Universal Robots URScript: letra_E.script

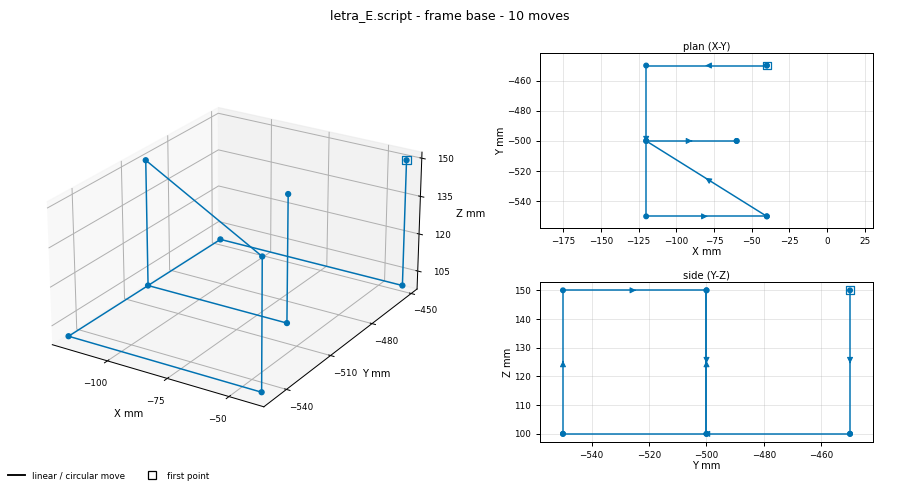
[picture p0: tool path of letra_E.script in frame base, 10 of 10 moves have a stored position in this frame; points joined in program order, loops and branches not executed]
# Letra E - Escobar
movel(p[-0.040, -0.450, 0.150, 3.1416, 0, 0], a=0.5, v=0.1)
movel(p[-0.040, -0.450, 0.100, 3.1416, 0, 0], a=0.5, v=0.1)
movel(p[-0.120, -0.450, 0.100, 3.1416, 0, 0], a=0.5, v=0.1)
movel(p[-0.120, -0.550, 0.100, 3.1416, 0, 0], a=0.5, v=0.1)
movel(p[-0.040, -0.550, 0.100, 3.1416, 0, 0], a=0.5, v=0.1)
movel(p[-0.040, -0.550, 0.150, 3.1416, 0, 0], a=0.5, v=0.1)
movel(p[-0.120, -0.500, 0.150, 3.1416, 0, 0], a=0.5, v=0.1)
movel(p[-0.120, -0.500, 0.100, 3.1416, 0, 0], a=0.5, v=0.1)
movel(p[-0.060, -0.500, 0.100, 3.1416, 0, 0], a=0.5, v=0.1)
movel(p[-0.060, -0.500, 0.150, 3.1416, 0, 0], a=0.5, v=0.1)
